Fanuc KAREL source: kb00018.KL

-- PROVISIONAL review KL for V940-1; original PC SHA256 ab2243a005f9ca8637fba59ff8659a50f60370f0190641cda7dbfd95330b134a
-- Incomplete behavior may be omitted. Consult companion uncertainty JSON. Do not deploy.
PROGRAM KB00018
%NOLOCKGROUP
BEGIN
  -- V9_ZERO_TABLE_METADATA_HINT layout=0002_ascii; no indexed target words; source/name/runtime held
  -- UNRESOLVED_PC offsets 5-12; opcodes 9D,23
  -- UNRESOLVED_PC offsets 17-65; opcodes 27,22,1C,22,1C,22,1C,22,27,9D,31
  -- UNRESOLVED_PC offsets 70-74; opcodes 7F
END KB00018
